FUNCTION_BLOCK MOD_ActivityCount (* Counts the skills that are running: every skill says +1 when it starts and -1 when it ends. Technical: Number of running skills from the +1/-1 activity channel *)
  (* Standard: 61499-2 *)
  (* Version 0.1, 2026-09-28, Project contributors, AAU Smart Production Lab *)
  PACKAGE modlib;
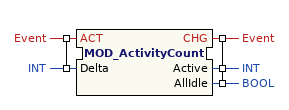
  EVENT_INPUT
    ACT WITH Delta; (* A skill started (+1) or ended (-1) *)
  END_EVENT
  EVENT_OUTPUT
    CHG WITH Active, AllIdle; (* The value changed *)
  END_EVENT
  VAR_INPUT
    Delta : INT; (* +1 when a skill starts, -1 when it ends *)
  END_VAR
  VAR_OUTPUT
    Active : INT; (* Some skill runs *)
    AllIdle : BOOL := TRUE; (* No skill runs *)
  END_VAR
  EC_STATES
    ACT : ACT -> CHG;
  END_STATES
  ALGORITHM ACT IN ST:
Active := Active + Delta;
IF Active < 0 THEN
  Active := 0;
END_IF;
AllIdle := Active = 0;
  END_ALGORITHM
END_FUNCTION_BLOCK
